// TIA Portal V20 export
Screen "Robot_Kuka"  1276x673
  ScreenItem "permanentareaborderrectangle" at 0,0 size 0x0  Type=HmiRectangle
  ScreenItem "Line_Header_X0_Y64" at 0,64 size 1276x0  Type=HmiLine
  ScreenItem "Select Robot" at 487,68 size 290x37  Type=HmiSymbolicIOField
  ScreenItem "Button_Back" at 2,2 size 90x60  Type=HmiButton
  ScreenItem "Button_Collision" at 93,2 size 90x60  Type=HmiButton
  ScreenItem "Title_ScreenOverview_X390_Y2_3" at 252,816 size 497x59  Type=HmiTextBox
  ScreenItem "Robot Name" at 275,816 size 192x52  Type=HmiIOField
  ScreenItem "Button_Collision_3" at 1253,802 size 90x60  Type=HmiButton
  ScreenItem "Button_Collision_6" at 1253,802 size 90x60  Type=HmiButton
  ScreenItem "140RB03" at 0,0 size 90x60  Type=HmiButton
  ScreenItem "140RB01_5" at 0,0 size 90x60  Type=HmiButton
  ScreenItem "140RB01_1" at 0,0 size 90x60  Type=HmiButton
  ScreenItem "140RB01_2" at 0,0 size 90x60  Type=HmiButton
  ScreenItem "140RB01_3" at 0,0 size 90x60  Type=HmiButton
  ScreenItem "140RB01_4" at 0,0 size 90x60  Type=HmiButton
  ScreenItem "Select Robot_1" at 398,8 size 473x48  Type=HmiSymbolicIOField
  ScreenItem "矩形_50" at 0,0 size 328x297  Type=HmiRectangle
  ScreenItem "矩形_1" at 31,47 size 17x17  Type=HmiRectangle
  ScreenItem "文本_1" at 56,26 size 39x22  Type=HmiText
  ScreenItem "文本_2" at 20,26 size 39x22  Type=HmiText
  ScreenItem "矩形_2" at 63,47 size 17x17  Type=HmiRectangle
  ScreenItem "文本_3" at 11,47 size 16x17  Type=HmiText
  ScreenItem "文本_4" at 11,67 size 16x17  Type=HmiText
  ScreenItem "文本_5" at 11,87 size 16x17  Type=HmiText
  ScreenItem "文本_6" at 11,107 size 16x17  Type=HmiText
  ScreenItem "文本_7" at 11,127 size 16x17  Type=HmiText
  ScreenItem "文本_8" at 11,147 size 16x17  Type=HmiText
  ScreenItem "文本_9" at 11,167 size 16x17  Type=HmiText
  ScreenItem "文本_10" at 11,187 size 16x17  Type=HmiText
  ScreenItem "文本_11" at 11,207 size 16x17  Type=HmiText
  ScreenItem "文本_12" at 11,227 size 16x17  Type=HmiText
  ScreenItem "文本_13" at 11,247 size 16x17  Type=HmiText
  ScreenItem "文本_14" at 12,267 size 15x17  Type=HmiText
  ScreenItem "文本_15" at 139,26 size 39x22  Type=HmiText
  ScreenItem "文本_16" at 109,26 size 39x22  Type=HmiText
  ScreenItem "文本_17" at 100,47 size 16x17  Type=HmiText
  ScreenItem "文本_18" at 100,67 size 16x17  Type=HmiText
  ScreenItem "文本_19" at 100,87 size 16x17  Type=HmiText
  ScreenItem "文本_20" at 100,107 size 16x17  Type=HmiText
  ScreenItem "文本_21" at 100,127 size 16x17  Type=HmiText
  ScreenItem "文本_22" at 100,147 size 16x17  Type=HmiText
  ScreenItem "文本_23" at 100,167 size 16x17  Type=HmiText
  ScreenItem "文本_24" at 100,187 size 16x17  Type=HmiText
  ScreenItem "文本_25" at 100,207 size 16x17  Type=HmiText
  ScreenItem "文本_26" at 100,227 size 16x17  Type=HmiText
  ScreenItem "文本_27" at 100,247 size 16x17  Type=HmiText
  ScreenItem "文本_28" at 100,267 size 16x17  Type=HmiText
  ScreenItem "文本_29" at 198,47 size 16x17  Type=HmiText
  ScreenItem "文本_30" at 198,69 size 16x17  Type=HmiText
  ScreenItem "文本_31" at 198,89 size 16x17  Type=HmiText
  ScreenItem "文本_32" at 198,109 size 16x17  Type=HmiText
  ScreenItem "文本_33" at 271,47 size 16x16  Type=HmiText
  ScreenItem "文本_34" at 271,69 size 16x17  Type=HmiText
  ScreenItem "文本_35" at 271,89 size 16x17  Type=HmiText
  ScreenItem "文本_36" at 198,206 size 16x17  Type=HmiText
  ScreenItem "文本_37" at 198,226 size 16x17  Type=HmiText
  ScreenItem "文本_38" at 198,246 size 16x17  Type=HmiText
  ScreenItem "文本_39" at 198,266 size 16x17  Type=HmiText
  ScreenItem "Text field_DoDockRel1_1" at 9,0 size 171x27  Type=HmiTextBox
  ScreenItem "线_1" at 187,0 size 0x298  Type=HmiLine
  ScreenItem "Text field_DoDockRel1_2" at 196,1 size 124x27  Type=HmiTextBox
  ScreenItem "Text field_DoDockRel1_3" at 197,143 size 124x48  Type=HmiTextBox
  ScreenItem "矩形_52" at 31,67 size 17x17  Type=HmiRectangle
  ScreenItem "矩形_3" at 31,87 size 17x17  Type=HmiRectangle
  ScreenItem "矩形_4" at 31,107 size 17x17  Type=HmiRectangle
  ScreenItem "矩形_5" at 31,127 size 17x17  Type=HmiRectangle
  ScreenItem "矩形_7" at 31,147 size 17x17  Type=HmiRectangle
  ScreenItem "矩形_9" at 31,167 size 17x17  Type=HmiRectangle
  ScreenItem "矩形_11" at 31,187 size 17x17  Type=HmiRectangle
  ScreenItem "矩形_13" at 31,207 size 17x17  Type=HmiRectangle
  ScreenItem "矩形_15" at 31,227 size 17x17  Type=HmiRectangle
  ScreenItem "矩形_17" at 31,247 size 17x17  Type=HmiRectangle
  ScreenItem "矩形_19" at 31,267 size 17x17  Type=HmiRectangle
  ScreenItem "矩形_6" at 63,67 size 17x17  Type=HmiRectangle
  ScreenItem "矩形_8" at 63,87 size 17x17  Type=HmiRectangle
  ScreenItem "矩形_10" at 63,107 size 17x17  Type=HmiRectangle
  ScreenItem "矩形_12" at 63,127 size 17x17  Type=HmiRectangle
  ScreenItem "矩形_14" at 63,147 size 17x17  Type=HmiRectangle
  ScreenItem "矩形_16" at 63,167 size 17x17  Type=HmiRectangle
  ScreenItem "矩形_18" at 63,187 size 17x17  Type=HmiRectangle
  ScreenItem "矩形_20" at 63,207 size 17x17  Type=HmiRectangle
  ScreenItem "矩形_21" at 63,227 size 17x17  Type=HmiRectangle
  ScreenItem "矩形_22" at 63,247 size 17x17  Type=HmiRectangle
  ScreenItem "矩形_23" at 63,267 size 17x17  Type=HmiRectangle
  ScreenItem "矩形_24" at 122,47 size 17x17  Type=HmiRectangle
  ScreenItem "矩形_25" at 152,47 size 17x17  Type=HmiRectangle
  ScreenItem "矩形_26" at 122,66 size 17x17  Type=HmiRectangle
  ScreenItem "矩形_27" at 122,86 size 17x17  Type=HmiRectangle
  ScreenItem "矩形_28" at 122,106 size 17x17  Type=HmiRectangle
  ScreenItem "矩形_29" at 122,126 size 17x17  Type=HmiRectangle
  ScreenItem "矩形_30" at 122,146 size 17x17  Type=HmiRectangle
  ScreenItem "矩形_31" at 122,166 size 17x17  Type=HmiRectangle
  ScreenItem "矩形_32" at 122,186 size 17x17  Type=HmiRectangle
  ScreenItem "矩形_33" at 122,206 size 17x17  Type=HmiRectangle
  ScreenItem "矩形_34" at 122,226 size 17x17  Type=HmiRectangle
  ScreenItem "矩形_35" at 122,246 size 17x17  Type=HmiRectangle
  ScreenItem "矩形_36" at 122,266 size 17x17  Type=HmiRectangle
  ScreenItem "矩形_37" at 152,66 size 17x17  Type=HmiRectangle
  ScreenItem "矩形_38" at 152,86 size 17x17  Type=HmiRectangle
  ScreenItem "矩形_39" at 152,106 size 17x17  Type=HmiRectangle
  ScreenItem "矩形_40" at 152,126 size 17x17  Type=HmiRectangle
  ScreenItem "矩形_41" at 152,146 size 17x17  Type=HmiRectangle
  ScreenItem "矩形_42" at 152,166 size 17x17  Type=HmiRectangle
  ScreenItem "矩形_43" at 152,186 size 17x17  Type=HmiRectangle
  ScreenItem "矩形_44" at 152,206 size 17x17  Type=HmiRectangle
  ScreenItem "矩形_45" at 152,226 size 17x17  Type=HmiRectangle
  ScreenItem "矩形_46" at 152,246 size 17x17  Type=HmiRectangle
  ScreenItem "矩形_47" at 152,266 size 17x17  Type=HmiRectangle
  ScreenItem "矩形_48" at 213,47 size 17x17  Type=HmiRectangle
  ScreenItem "矩形_49" at 213,68 size 17x17  Type=HmiRectangle
  ScreenItem "矩形_51" at 213,88 size 17x17  Type=HmiRectangle
  ScreenItem "矩形_53" at 213,108 size 17x17  Type=HmiRectangle
  ScreenItem "矩形_54" at 287,47 size 17x17  Type=HmiRectangle
  ScreenItem "矩形_55" at 287,68 size 17x17  Type=HmiRectangle
  ScreenItem "矩形_56" at 287,88 size 17x17  Type=HmiRectangle
  ScreenItem "矩形_57" at 213,206 size 17x17  Type=HmiRectangle
  ScreenItem "矩形_58" at 213,226 size 17x17  Type=HmiRectangle
  ScreenItem "矩形_59" at 213,246 size 17x17  Type=HmiRectangle
  ScreenItem "矩形_60" at 213,266 size 17x17  Type=HmiRectangle
  ScreenItem "acABBMessages" at 735,125 size 528x522  Type=HmiAlarmControl
  ScreenItem "Rectangle Segment Status" at 303,125 size 284x520  Type=HmiRectangle
  ScreenItem "Rectangle Robot Status" at 19,125 size 284x394  Type=HmiRectangle
  ScreenItem "Text Filed E- Stop" at 160,228 size 128x21  Type=HmiTextBox
  ScreenItem "Text Field In Auto On" at 25,159 size 128x21  Type=HmiTextBox
  ScreenItem "Text Field Home Position" at 25,182 size 128x21  Type=HmiTextBox
  ScreenItem "Text field Robot Status" at 19,124 size 284x31  Type=HmiTextBox
  ScreenItem "Rectangle Collision Zone" at 19,520 size 283x125  Type=HmiRectangle
  ScreenItem "ClearZone1" at 24,552 size 31x20  Type=HmiRectangle
  ScreenItem "ReqZone1" at 24,552 size 31x20  Type=HmiRectangle
  ScreenItem "Fault_1" at 24,552 size 31x20  Type=HmiRectangle
  ScreenItem "TextZone1" at 24,552 size 31x20  Type=HmiText
  ScreenItem "ClearZone2" at 59,552 size 31x20  Type=HmiRectangle
  ScreenItem "ReqZone2" at 59,552 size 31x20  Type=HmiRectangle
  ScreenItem "Fault_2" at 59,552 size 31x20  Type=HmiRectangle
  ScreenItem "TextZone2" at 59,552 size 31x20  Type=HmiText
  ScreenItem "ClearZone3" at 93,552 size 31x20  Type=HmiRectangle
  ScreenItem "ReqZone3" at 93,552 size 31x20  Type=HmiRectangle
  ScreenItem "Fault_3" at 93,552 size 31x20  Type=HmiRectangle
  ScreenItem "TextZone3" at 93,552 size 31x20  Type=HmiText
  ScreenItem "ClearZone4" at 128,552 size 31x20  Type=HmiRectangle
  ScreenItem "ReqZone4" at 128,552 size 31x20  Type=HmiRectangle
  ScreenItem "Fault_4" at 128,552 size 31x20  Type=HmiRectangle
  ScreenItem "TextZone4" at 128,552 size 31x20  Type=HmiText
  ScreenItem "ClearZone5" at 162,552 size 31x20  Type=HmiRectangle
  ScreenItem "ReqZone5" at 162,552 size 31x20  Type=HmiRectangle
  ScreenItem "Fault_5" at 162,552 size 31x20  Type=HmiRectangle
  ScreenItem "TextZone5" at 162,552 size 31x20  Type=HmiText
  ScreenItem "ClearZone6" at 197,552 size 31x20  Type=HmiRectangle
  ScreenItem "ReqZone6" at 197,552 size 31x20  Type=HmiRectangle
  ScreenItem "Fault_6" at 197,552 size 31x20  Type=HmiRectangle
  ScreenItem "TextZone6" at 197,552 size 31x20  Type=HmiText
  ScreenItem "ClearZone7" at 232,552 size 31x20  Type=HmiRectangle
  ScreenItem "ReqZone7" at 232,552 size 31x20  Type=HmiRectangle
  ScreenItem "Fault_7" at 232,552 size 31x20  Type=HmiRectangle
  ScreenItem "TextZone7" at 232,552 size 31x20  Type=HmiText
  ScreenItem "ClearZone8" at 266,552 size 31x20  Type=HmiRectangle
  ScreenItem "ReqZone8" at 266,552 size 31x20  Type=HmiRectangle
  ScreenItem "Fault_8" at 266,552 size 31x20  Type=HmiRectangle
  ScreenItem "TextZone8" at 266,552 size 31x20  Type=HmiText
  ScreenItem "ClearZone9" at 24,575 size 31x20  Type=HmiRectangle
  ScreenItem "ReqZone9" at 24,575 size 31x20  Type=HmiRectangle
  ScreenItem "Fault_9" at 24,575 size 31x20  Type=HmiRectangle
  ScreenItem "TextZone9" at 24,575 size 31x20  Type=HmiText
  ScreenItem "ClearZone10" at 59,575 size 31x20  Type=HmiRectangle
  ScreenItem "ReqZone10" at 59,575 size 31x20  Type=HmiRectangle
  ScreenItem "Fault_10" at 59,575 size 31x20  Type=HmiRectangle
  ScreenItem "TextZone10" at 59,575 size 31x20  Type=HmiText
  ScreenItem "ClearZone11" at 93,575 size 31x20  Type=HmiRectangle
  ScreenItem "ReqZone11" at 93,575 size 31x20  Type=HmiRectangle
  ScreenItem "Fault_11" at 93,575 size 31x20  Type=HmiRectangle
  ScreenItem "TextZone11" at 93,575 size 31x20  Type=HmiText
  ScreenItem "ClearZone12" at 128,575 size 31x20  Type=HmiRectangle
  ScreenItem "ReqZone12" at 128,575 size 31x20  Type=HmiRectangle
  ScreenItem "Fault_12" at 128,575 size 31x20  Type=HmiRectangle
  ScreenItem "TextZone12" at 128,575 size 31x20  Type=HmiText
  ScreenItem "ClearZone13" at 162,575 size 31x20  Type=HmiRectangle
  ScreenItem "ReqZone13" at 162,575 size 31x20  Type=HmiRectangle
  ScreenItem "Fault_13" at 162,575 size 31x20  Type=HmiRectangle
  ScreenItem "TextZone13" at 162,575 size 31x20  Type=HmiText
  ScreenItem "ClearZone14" at 197,575 size 31x20  Type=HmiRectangle
  ScreenItem "ReqZone14" at 197,575 size 31x20  Type=HmiRectangle
  ScreenItem "Fault_14" at 197,575 size 31x20  Type=HmiRectangle
  ScreenItem "TextZone14" at 197,575 size 31x20  Type=HmiText
  ScreenItem "ClearZone15" at 232,575 size 31x20  Type=HmiRectangle
  ScreenItem "ReqZone15" at 232,575 size 31x20  Type=HmiRectangle
  ScreenItem "Fault_15" at 232,575 size 31x20  Type=HmiRectangle
  ScreenItem "TextZone15" at 232,575 size 31x20  Type=HmiText
  ScreenItem "ClearZone16" at 266,575 size 31x20  Type=HmiRectangle
  ScreenItem "ReqZone16" at 266,575 size 31x20  Type=HmiRectangle
  ScreenItem "Fault_16" at 266,575 size 31x20  Type=HmiRectangle
  ScreenItem "TextZone16" at 266,575 size 31x20  Type=HmiText
  ScreenItem "ClearZone17" at 24,598 size 31x20  Type=HmiRectangle
  ScreenItem "ReqZone17" at 24,598 size 31x20  Type=HmiRectangle
  ScreenItem "Fault_17" at 24,598 size 31x20  Type=HmiRectangle
  ScreenItem "TextZone17" at 24,598 size 31x20  Type=HmiText
  ScreenItem "ClearZone18" at 59,598 size 31x20  Type=HmiRectangle
  ScreenItem "ReqZone18" at 59,598 size 31x20  Type=HmiRectangle
  ScreenItem "Fault_18" at 59,598 size 31x20  Type=HmiRectangle
  ScreenItem "TextZone18" at 59,598 size 31x20  Type=HmiText
  ScreenItem "ClearZone19" at 93,598 size 31x20  Type=HmiRectangle
  ScreenItem "ReqZone19" at 93,598 size 31x20  Type=HmiRectangle
  ScreenItem "Fault_19" at 93,598 size 31x20  Type=HmiRectangle
  ScreenItem "TextZone19" at 93,598 size 31x20  Type=HmiText
  ScreenItem "ClearZone20" at 128,598 size 31x20  Type=HmiRectangle
  ScreenItem "ReqZone20" at 128,598 size 31x20  Type=HmiRectangle
  ScreenItem "Fault_20" at 128,598 size 31x20  Type=HmiRectangle
  ScreenItem "TextZone20" at 128,598 size 31x20  Type=HmiText
  ScreenItem "ClearZone21" at 162,598 size 31x20  Type=HmiRectangle
  ScreenItem "ReqZone21" at 162,598 size 31x20  Type=HmiRectangle
  ScreenItem "Fault_21" at 162,598 size 31x20  Type=HmiRectangle
  ScreenItem "TextZone21" at 162,598 size 31x20  Type=HmiText
  ScreenItem "ClearZone22" at 197,598 size 31x20  Type=HmiRectangle
  ScreenItem "ReqZone22" at 197,598 size 31x20  Type=HmiRectangle
  ScreenItem "Fault_22" at 197,598 size 31x20  Type=HmiRectangle
  ScreenItem "TextZone22" at 197,598 size 31x20  Type=HmiText
  ScreenItem "ClearZone23" at 232,598 size 31x20  Type=HmiRectangle
  ScreenItem "ReqZone23" at 232,598 size 31x20  Type=HmiRectangle
  ScreenItem "Fault_23" at 232,598 size 31x20  Type=HmiRectangle
  ScreenItem "TextZone23" at 232,598 size 31x20  Type=HmiText
  ScreenItem "ClearZone24" at 266,598 size 31x20  Type=HmiRectangle
  ScreenItem "ReqZone24" at 266,598 size 31x20  Type=HmiRectangle
  ScreenItem "Fault_24" at 266,598 size 31x20  Type=HmiRectangle
  ScreenItem "TextZone24" at 266,598 size 31x20  Type=HmiText
  ScreenItem "ClearZone25" at 24,621 size 31x20  Type=HmiRectangle
  ScreenItem "ReqZone25" at 24,621 size 31x20  Type=HmiRectangle
  ScreenItem "Fault_25" at 24,621 size 31x20  Type=HmiRectangle
  ScreenItem "TextZone25" at 24,621 size 31x20  Type=HmiText
  ScreenItem "ClearZone26" at 59,621 size 31x20  Type=HmiRectangle
  ScreenItem "ReqZone26" at 59,621 size 31x20  Type=HmiRectangle
  ScreenItem "Fault_26" at 59,621 size 31x20  Type=HmiRectangle
  ScreenItem "TextZone26" at 59,621 size 31x20  Type=HmiText
  ScreenItem "ClearZone27" at 93,621 size 31x20  Type=HmiRectangle
  ScreenItem "ReqZone27" at 93,621 size 31x20  Type=HmiRectangle
  ScreenItem "Fault_27" at 93,621 size 31x20  Type=HmiRectangle
  ScreenItem "TextZone27" at 93,621 size 31x20  Type=HmiText
  ScreenItem "ClearZone28" at 128,621 size 31x20  Type=HmiRectangle
  ScreenItem "ReqZone28" at 128,621 size 31x20  Type=HmiRectangle
  ScreenItem "Fault_28" at 128,621 size 31x20  Type=HmiRectangle
  ScreenItem "TextZone28" at 128,621 size 31x20  Type=HmiText
  ScreenItem "ClearZone29" at 162,621 size 31x20  Type=HmiRectangle
  ScreenItem "ReqZone29" at 162,621 size 31x20  Type=HmiRectangle
  ScreenItem "Fault_29" at 162,621 size 31x20  Type=HmiRectangle
  ScreenItem "TextZone29" at 162,621 size 31x20  Type=HmiText
  ScreenItem "ClearZone30" at 197,621 size 31x20  Type=HmiRectangle
  ScreenItem "ReqZone30" at 197,621 size 31x20  Type=HmiRectangle
  ScreenItem "Fault_30" at 197,621 size 31x20  Type=HmiRectangle
  ScreenItem "TextZone30" at 197,621 size 31x20  Type=HmiText
  ScreenItem "ClearZone31" at 232,621 size 31x20  Type=HmiRectangle
  ScreenItem "ReqZone31" at 232,621 size 31x20  Type=HmiRectangle
  ScreenItem "Fault_31" at 232,621 size 31x20  Type=HmiRectangle
  ScreenItem "TextZone31" at 232,621 size 31x20  Type=HmiText
  ScreenItem "ClearZone32" at 266,621 size 31x20  Type=HmiRectangle
  ScreenItem "ReqZone32" at 266,621 size 31x20  Type=HmiRectangle
  ScreenItem "Fault_32" at 266,621 size 31x20  Type=HmiRectangle
  ScreenItem "TextZone32" at 266,621 size 31x20  Type=HmiText
  ScreenItem "Text field Robot Collision Zone" at 19,519 size 284x31  Type=HmiTextBox
  ScreenItem "Text Field Manual" at 160,159 size 128x21  Type=HmiTextBox
  ScreenItem "Text Field System Ready" at 25,205 size 128x21  Type=HmiTextBox
  ScreenItem "Text Field Motor On" at 25,228 size 128x21  Type=HmiTextBox
  ScreenItem "Text Field In Cycle" at 25,251 size 128x21  Type=HmiTextBox
  ScreenItem "Text Field Cycle On" at 25,274 size 128x21  Type=HmiTextBox
  ScreenItem "Text Field On Path" at 25,297 size 128x21  Type=HmiTextBox
  ScreenItem "Text Field ProgNumReq" at 25,320 size 128x21  Type=HmiTextBox
  ScreenItem "Text Field Task OK" at 25,343 size 128x21  Type=HmiTextBox
  ScreenItem "Text Field Tryout Mode" at 160,182 size 128x21  Type=HmiTextBox
  ScreenItem "Text Field Stop" at 160,205 size 128x21  Type=HmiTextBox
  ScreenItem "Text Filed Error" at 160,251 size 128x21  Type=HmiTextBox
  ScreenItem "IO Field Feedback Program" at 160,369 size 128x21  Type=HmiIOField
  ScreenItem "Text Field Feedback Program" at 160,341 size 114x30  Type=HmiTextBox
  ScreenItem "Text Filed Process Fault" at 160,274 size 128x21  Type=HmiTextBox
  ScreenItem "Text field_DoOutSeg1" at 310,159 size 128x21  Type=HmiTextBox
  ScreenItem "Text field_DoOutSeg2" at 310,179 size 128x21  Type=HmiTextBox
  ScreenItem "Text field_DoOutSeg3" at 310,199 size 128x21  Type=HmiTextBox
  ScreenItem "Text field_DoOutSeg4" at 310,219 size 128x21  Type=HmiTextBox
  ScreenItem "Text field_DoOutSeg5" at 310,239 size 128x21  Type=HmiTextBox
  ScreenItem "Text field_DoOutSeg6" at 310,259 size 128x21  Type=HmiTextBox
  ScreenItem "Text field_DoOutSeg7" at 310,279 size 128x21  Type=HmiTextBox
  ScreenItem "Text field_DoOutSeg8" at 310,299 size 128x21  Type=HmiTextBox
  ScreenItem "Text field_DoOutSeg9" at 310,319 size 128x21  Type=HmiTextBox
  ScreenItem "Text field_DoOutSeg10" at 310,339 size 128x21  Type=HmiTextBox
  ScreenItem "Text field_DoOutSeg11" at 310,359 size 128x21  Type=HmiTextBox
  ScreenItem "Text field_DoOutSeg12" at 310,379 size 128x21  Type=HmiTextBox
  ScreenItem "Text field_DoOutSeg13" at 310,399 size 128x21  Type=HmiTextBox
  ScreenItem "Text field_DoOutSeg14" at 310,419 size 128x21  Type=HmiTextBox
  ScreenItem "Text field_DoOutSeg15" at 310,439 size 128x21  Type=HmiTextBox
  ScreenItem "Text field_DoOutSeg16" at 310,459 size 128x21  Type=HmiTextBox
  ScreenItem "Text field_DoOutSeg17" at 310,479 size 128x21  Type=HmiTextBox
  ScreenItem "Text field_DoOutSeg18" at 310,499 size 128x21  Type=HmiTextBox
  ScreenItem "Text field_DoOutSeg19" at 310,519 size 128x21  Type=HmiTextBox
  ScreenItem "Text field_DoOutSeg20" at 310,539 size 128x21  Type=HmiTextBox
  ScreenItem "Text field_DoOutSeg21" at 310,559 size 128x21  Type=HmiTextBox
  ScreenItem "Text field_DoOutSeg22" at 310,579 size 128x21  Type=HmiTextBox
  ScreenItem "Text field_DoOutSeg23" at 310,599 size 128x21  Type=HmiTextBox
  ScreenItem "Text field_DoOutSeg24" at 310,619 size 128x21  Type=HmiTextBox
  ScreenItem "Text field_DoFinishSeg1" at 444,159 size 128x21  Type=HmiTextBox
  ScreenItem "Text field_DoFinishSeg2" at 444,179 size 128x21  Type=HmiTextBox
  ScreenItem "Text field_DoFinishSeg3" at 444,199 size 128x21  Type=HmiTextBox
  ScreenItem "Text field_DoFinishSeg4" at 444,219 size 128x21  Type=HmiTextBox
  ScreenItem "Text field_DoFinishSeg5" at 444,239 size 128x21  Type=HmiTextBox
  ScreenItem "Text field_DoFinishSeg6" at 444,259 size 128x21  Type=HmiTextBox
  ScreenItem "Text field_DoFinishSeg7" at 444,279 size 128x21  Type=HmiTextBox
  ScreenItem "Text field_DoFinishSeg8" at 444,299 size 128x21  Type=HmiTextBox
  ScreenItem "Text field_DoFinishSeg9" at 444,319 size 128x21  Type=HmiTextBox
  ScreenItem "Text field_DoFinishSeg10" at 444,339 size 128x21  Type=HmiTextBox
  ScreenItem "Text field_DoFinishSeg11" at 444,359 size 128x21  Type=HmiTextBox
  ScreenItem "Text field_DoFinishSeg12" at 444,379 size 128x21  Type=HmiTextBox
  ScreenItem "Text field_DoFinishSeg13" at 444,399 size 128x21  Type=HmiTextBox
  ScreenItem "Text field_DoFinishSeg14" at 444,419 size 128x21  Type=HmiTextBox
  ScreenItem "Text field_DoFinishSeg15" at 444,439 size 128x21  Type=HmiTextBox
  ScreenItem "Text field_DoFinishSeg16" at 444,459 size 128x21  Type=HmiTextBox
  ScreenItem "Text field_DoFinishSeg17" at 444,479 size 128x21  Type=HmiTextBox
  ScreenItem "Text field_DoFinishSeg18" at 444,499 size 128x21  Type=HmiTextBox
  ScreenItem "Text field_DoFinishSeg19" at 444,519 size 128x21  Type=HmiTextBox
  ScreenItem "Text field_DoFinishSeg20" at 444,539 size 128x21  Type=HmiTextBox
  ScreenItem "Text field_DoFinishSeg21" at 444,559 size 128x21  Type=HmiTextBox
  ScreenItem "Text field_DoFinishSeg22" at 444,579 size 128x21  Type=HmiTextBox
  ScreenItem "Text field_DoFinishSeg23" at 444,599 size 128x21  Type=HmiTextBox
  ScreenItem "Text field_DoFinishSeg24" at 444,619 size 128x21  Type=HmiTextBox
  ScreenItem "Text field Segment Status" at 303,124 size 284x31  Type=HmiTextBox
  ScreenItem "Text field Weld Spot Count" at 19,403 size 284x31  Type=HmiTextBox
  ScreenItem "Rectangle Dock Status" at 588,125 size 147x520  Type=HmiRectangle
  ScreenItem "Text field Dock Status" at 588,124 size 147x31  Type=HmiTextBox
  ScreenItem "Text field_DoDockRel1" at 594,159 size 128x21  Type=HmiTextBox
  ScreenItem "Text field_DoDockRel2" at 594,205 size 128x21  Type=HmiTextBox
  ScreenItem "Text field_DoDockRel3" at 594,251 size 128x21  Type=HmiTextBox
  ScreenItem "Text field_DoDockRel4" at 594,297 size 128x21  Type=HmiTextBox
  ScreenItem "Text field_DoDockEnd1" at 594,179 size 128x21  Type=HmiTextBox
  ScreenItem "Text field_DoDockEnd2" at 594,225 size 128x21  Type=HmiTextBox
  ScreenItem "Text field_DoDockEnd3" at 594,271 size 128x21  Type=HmiTextBox
  ScreenItem "Text field_DoDockEnd4" at 594,317 size 128x21  Type=HmiTextBox
  ScreenItem "Text field World Zone" at 588,346 size 147x31  Type=HmiTextBox
  ScreenItem "Text field_DoWorldZone1" at 594,381 size 128x21  Type=HmiTextBox
  ScreenItem "Text field_DoWorldZone2" at 594,404 size 128x21  Type=HmiTextBox
  ScreenItem "Text field_DoWorldZone3" at 594,427 size 128x21  Type=HmiTextBox
  ScreenItem "Text field_DoWorldZone4" at 594,450 size 128x21  Type=HmiTextBox
  ScreenItem "Text field_DoWorldZone5" at 594,473 size 128x21  Type=HmiTextBox
  ScreenItem "Text field_DoWorldZone6" at 594,496 size 128x21  Type=HmiTextBox
  ScreenItem "Text field_DoWorldZone7" at 594,519 size 128x21  Type=HmiTextBox
  ScreenItem "Text field_DoWorldZone8" at 594,542 size 128x21  Type=HmiTextBox
  ScreenItem "Text Field Home Position_1" at 160,297 size 128x21  Type=HmiTextBox
  ScreenItem "Text Field Home Position_2" at 160,320 size 128x21  Type=HmiTextBox
  ScreenItem "Text Field Feedback Program_1" at 31,357 size 114x30  Type=HmiTextBox
  ScreenItem "IO Field Feedback Program_1" at 27,379 size 128x21  Type=HmiIOField
  ScreenItem "Text Field WeldSpotCount" at 53,433 size 147x21  Type=HmiTextBox
  ScreenItem "IO Field Weld Spot Count" at 204,435 size 61x21  Type=HmiIOField
  ScreenItem "Rectangle Bypass Weld Count" at 180,460 size 85x55  Type=HmiRectangle
  ScreenItem "Button Bypass Weld Count" at 181,461 size 83x54  Type=HmiButton
  ScreenItem "Text Field WeldSpotCount_1" at 51,462 size 24x21  Type=HmiTextBox
  ScreenItem "IO Field Weld Spot Count_1" at 72,462 size 37x21  Type=HmiIOField
  ScreenItem "Text Field WeldSpotCount_2" at 116,462 size 24x21  Type=HmiTextBox
  ScreenItem "IO Field Weld Spot Count_2" at 137,462 size 37x21  Type=HmiIOField
  ScreenItem "Text Field WeldSpotCount_3" at 51,487 size 24x21  Type=HmiTextBox
  ScreenItem "IO Field Weld Spot Count_3" at 72,487 size 37x21  Type=HmiIOField
  ScreenItem "Text Field WeldSpotCount_4" at 116,487 size 24x21  Type=HmiTextBox
  ScreenItem "IO Field Weld Spot Count_4" at 137,487 size 37x21  Type=HmiIOField
  ScreenItem "Button_Collision_9" at 184,1 size 90x60  Type=HmiButton
